TYPE "FRK_PermCtx"
VERSION : 0.1
   STRUCT
      "Permit" : Bool;
      "Count" : Int;
      "Blocker" : String[160];
   END_STRUCT;
END_TYPE
